(* PLC project Vn_xor2, Beckhoff Automation GmbH TwinCAT PLC Control 3.5.13.21 *)
(* stored: creationDateTime 1970-01-01T00:00:00 *)

PROGRAM Vn_xor2

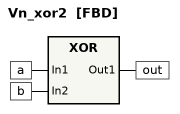
(* FBD diagram, written out as Structured Text *)
out := a XOR b;
END_PROGRAM
